ABB RAPID module: SpeedProg.mod

MODULE MainModule
GLOBAL VAR robtarget robpoint0= p:{{-607.850, 543.849, 363.215},{0.374108, 0.285846, 0.853660, -0.222712}}{cfg 0,0,0,0}{EJ 0.000000000,0.000000000,0.000000000,0.000000000,0.000000000,0.000000000}
GLOBAL VAR robtarget robpoint1= p:{{-640.584, 506.980, 371.534},{0.374108, 0.285846, 0.853660, -0.222712}}{cfg 0,0,0,0}{EJ 0.000000000,0.000000000,0.000000000,0.000000000,0.000000000,0.000000000}
GLOBAL VAR robtarget robpoint2= p:{{-607.850, 543.849, 363.215},{0.374108, 0.285846, 0.853660, -0.222712}}{cfg 0,0,0,0}{EJ 0.000000000,0.000000000,0.000000000,0.000000000,0.000000000,0.000000000}
GLOBAL VAR robtarget robpoint3= p:{{-640.584, 506.980, 371.534},{0.374108, 0.285846, 0.853660, -0.222712}}{cfg 0,0,0,0}{EJ 0.000000000,0.000000000,0.000000000,0.000000000,0.000000000,0.000000000}
GLOBAL VAR robtarget robpoint4= p:{{-607.850, 543.849, 363.215},{0.374108, 0.285846, 0.853660, -0.222712}}{cfg 0,0,0,0}{EJ 0.000000000,0.000000000,0.000000000,0.000000000,0.000000000,0.000000000}
GLOBAL VAR robtarget robpoint5= p:{{-640.584, 506.980, 371.534},{0.374108, 0.285846, 0.853660, -0.222712}}{cfg 0,0,0,0}{EJ 0.000000000,0.000000000,0.000000000,0.000000000,0.000000000,0.000000000}
GLOBAL VAR robtarget robpoint6= p:{{-607.850, 543.849, 363.215},{0.374108, 0.285846, 0.853660, -0.222712}}{cfg 0,0,0,0}{EJ 0.000000000,0.000000000,0.000000000,0.000000000,0.000000000,0.000000000}
GLOBAL VAR robtarget robpoint7= p:{{-640.584, 506.980, 371.534},{0.374108, 0.285846, 0.853660, -0.222712}}{cfg 0,0,0,0}{EJ 0.000000000,0.000000000,0.000000000,0.000000000,0.000000000,0.000000000}
GLOBAL VAR robtarget robpoint8= p:{{-607.850, 543.849, 363.215},{0.374108, 0.285846, 0.853660, -0.222712}}{cfg 0,0,0,0}{EJ 0.000000000,0.000000000,0.000000000,0.000000000,0.000000000,0.000000000}
GLOBAL VAR robtarget robpoint9= p:{{-640.584, 506.980, 371.534},{0.374108, 0.285846, 0.853660, -0.222712}}{cfg 0,0,0,0}{EJ 0.000000000,0.000000000,0.000000000,0.000000000,0.000000000,0.000000000}
GLOBAL VAR robtarget robpoint10= p:{{-640.584, 506.980, 371.534},{0.374108, 0.285846, 0.853660, -0.222712}}{cfg 0,0,0,0}{EJ 0.000000000,0.000000000,0.000000000,0.000000000,0.000000000,0.000000000}

GLOBAL Proc main()
    wobj16.x = 1234.57
    wobj16.y = -98.765
    wobj16.z = 50.500
    wobj16.q1 = 0.965926
    wobj16.q2 = 0.000000
    wobj16.q3 = 0.000000
    wobj16.q4 = 0.258819
    tool03.x = 10.000
    tool03.y = 20.000
    tool03.z = 150.000
    tool03.q1 = 1.000000
    tool03.q2 = 0.000000
    tool03.q3 = 0.000000
    tool03.q4 = 0.000000
    MoveL robpoint0,v1,z0,tool03,wobj16
    MoveL robpoint1,v12,z1,tool03,wobj16
    MoveL robpoint2,v99,z2,tool03,wobj16
    MoveL robpoint3,v333,z3,tool03,wobj16
    MoveL robpoint4,v1000,z6,tool03,wobj16
    MoveL robpoint5,v2500,z9,tool03,wobj16
    MoveL robpoint6,v5000,z15,tool03,wobj16
    MoveL robpoint7,v12000,z30,tool03,wobj16
    MoveL robpoint8,v0,z75,tool03,wobj16
    MoveL robpoint9,v750,z150,tool03,wobj16
    MoveL robpoint10,v750,z150,tool03,wobj16
EndProc
EndModule
